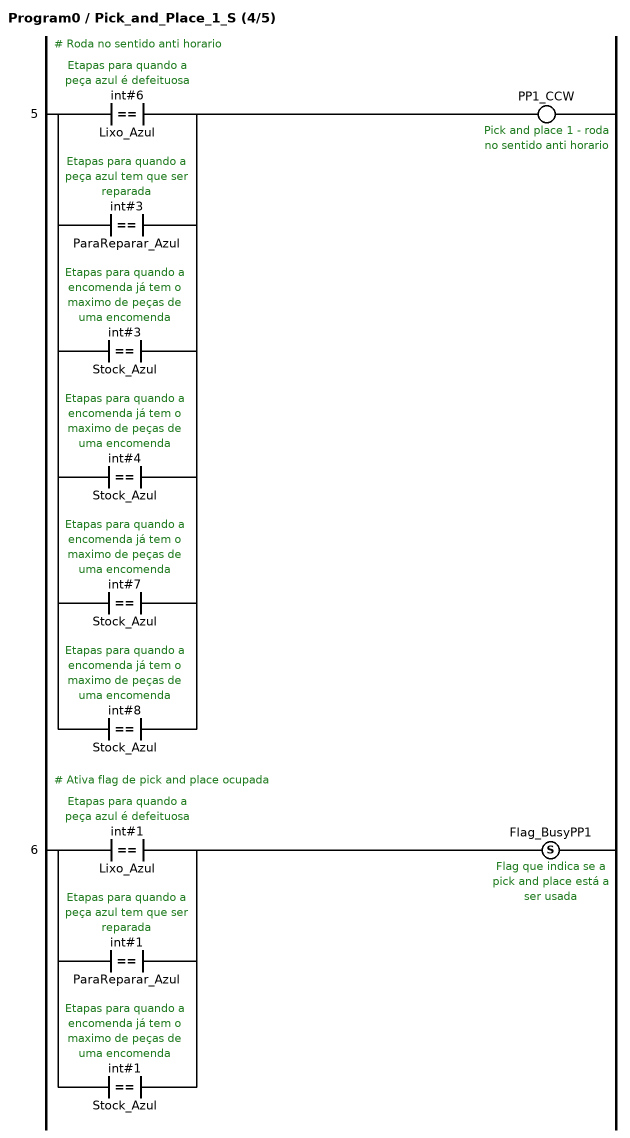
(* [picture p48: Program0 / Pick_and_Place_1_S, rungs 5-6] *)
(* Rung 5: # Roda no sentido anti horario *)
PP1_CCW := (int#6 = Lixo_Azul) OR (int#3 = ParaReparar_Azul) OR (int#3 = Stock_Azul) OR (int#4 = Stock_Azul) OR (int#7 = Stock_Azul) OR (int#8 = Stock_Azul);
(* Rung 6: # Ativa flag de pick and place ocupada *)
IF (int#1 = Lixo_Azul) OR (int#1 = ParaReparar_Azul) OR (int#1 = Stock_Azul) THEN
    Flag_BusyPP1 := TRUE;
END_IF;

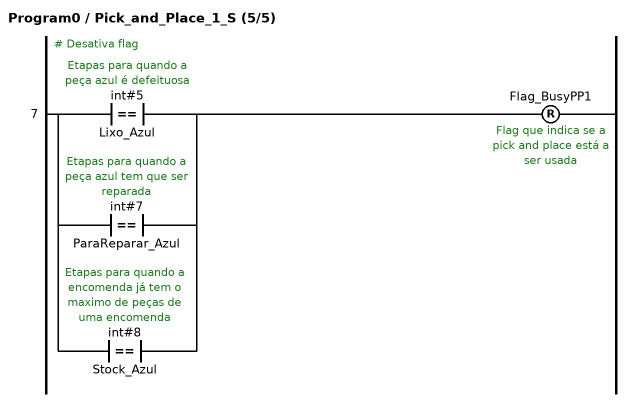
(* Rung 7: # Desativa flag *)
IF (int#5 = Lixo_Azul) OR (int#7 = ParaReparar_Azul) OR (int#8 = Stock_Azul) THEN
    Flag_BusyPP1 := FALSE;
END_IF;

(* Section Pick_and_Place_2_S: ladder, written here as Structured Text *)

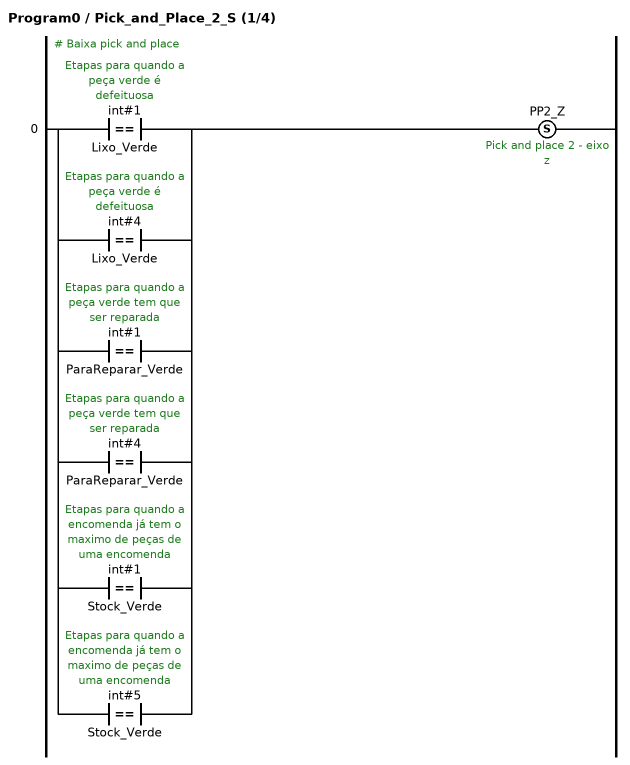
(* Rung 0: # Baixa pick and place *)
IF (int#1 = Lixo_Verde) OR (int#4 = Lixo_Verde) OR (int#1 = ParaReparar_Verde) OR (int#4 = ParaReparar_Verde) OR (int#1 = Stock_Verde) OR (int#5 = Stock_Verde) THEN
    PP2_Z := TRUE;
END_IF;

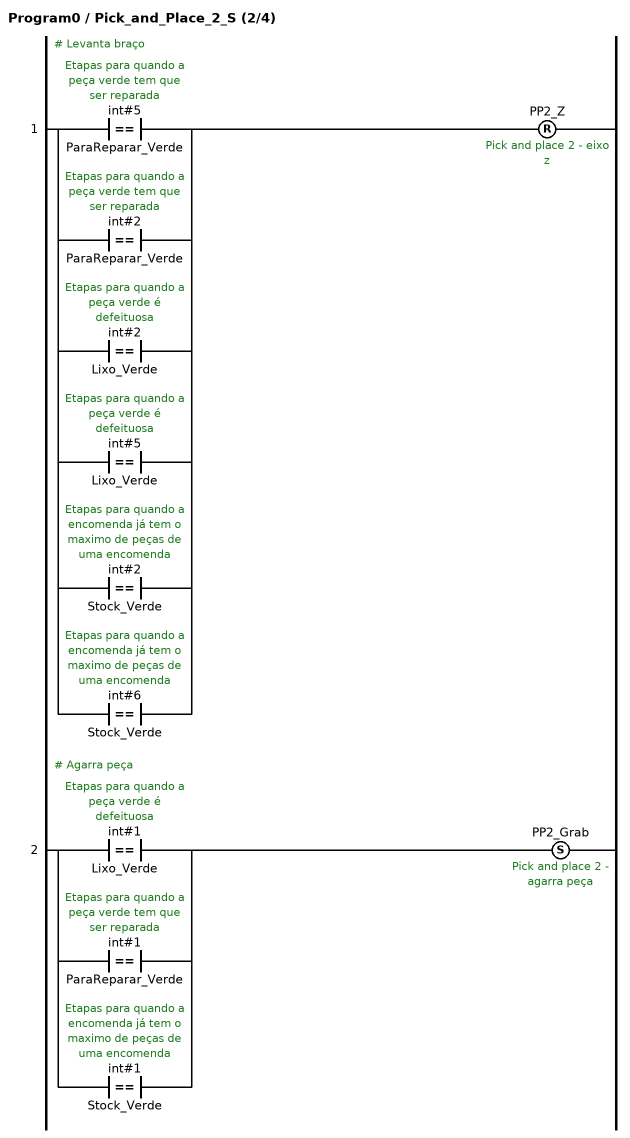
(* Rung 1: # Levanta braço *)
IF (int#5 = ParaReparar_Verde) OR (int#2 = ParaReparar_Verde) OR (int#2 = Lixo_Verde) OR (int#5 = Lixo_Verde) OR (int#2 = Stock_Verde) OR (int#6 = Stock_Verde) THEN
    PP2_Z := FALSE;
END_IF;
(* Rung 2: # Agarra peça *)
IF (int#1 = Lixo_Verde) OR (int#1 = ParaReparar_Verde) OR (int#1 = Stock_Verde) THEN
    PP2_Grab := TRUE;
END_IF;

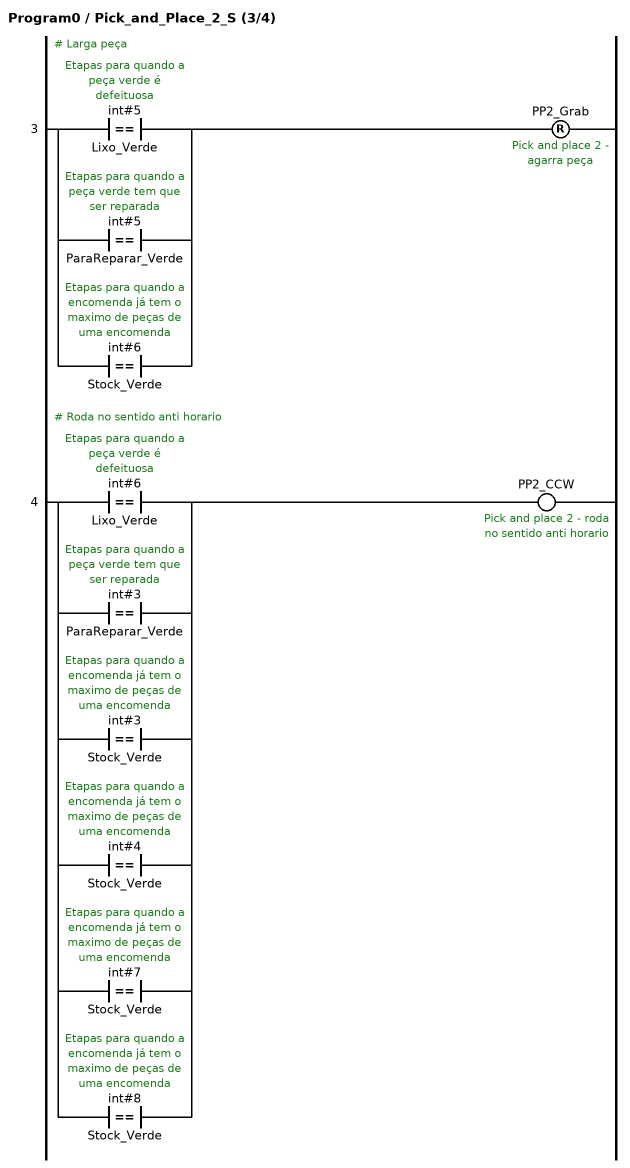
(* Rung 3: # Larga peça *)
IF (int#5 = Lixo_Verde) OR (int#5 = ParaReparar_Verde) OR (int#6 = Stock_Verde) THEN
    PP2_Grab := FALSE;
END_IF;
(* Rung 4: # Roda no sentido anti horario *)
PP2_CCW := (int#6 = Lixo_Verde) OR (int#3 = ParaReparar_Verde) OR (int#3 = Stock_Verde) OR (int#4 = Stock_Verde) OR (int#7 = Stock_Verde) OR (int#8 = Stock_Verde);

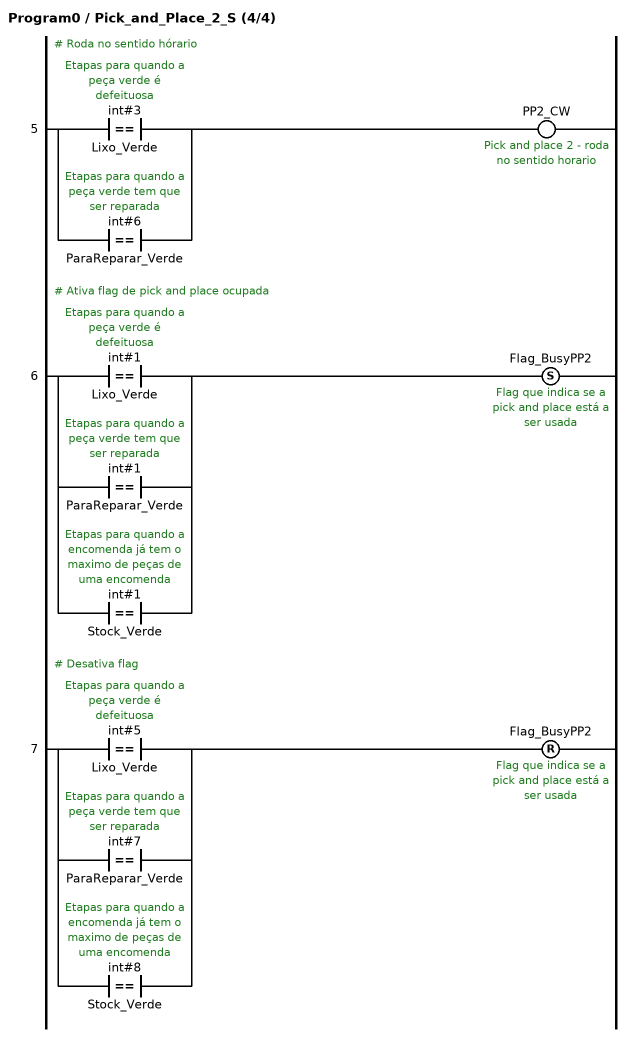
(* Rung 5: # Roda no sentido hórario *)
PP2_CW := (int#3 = Lixo_Verde) OR (int#6 = ParaReparar_Verde);
(* Rung 6: # Ativa flag de pick and place ocupada *)
IF (int#1 = Lixo_Verde) OR (int#1 = ParaReparar_Verde) OR (int#1 = Stock_Verde) THEN
    Flag_BusyPP2 := TRUE;
END_IF;
(* Rung 7: # Desativa flag *)
IF (int#5 = Lixo_Verde) OR (int#7 = ParaReparar_Verde) OR (int#8 = Stock_Verde) THEN
    Flag_BusyPP2 := FALSE;
END_IF;

(* Section Botoes: ladder, written here as Structured Text *)

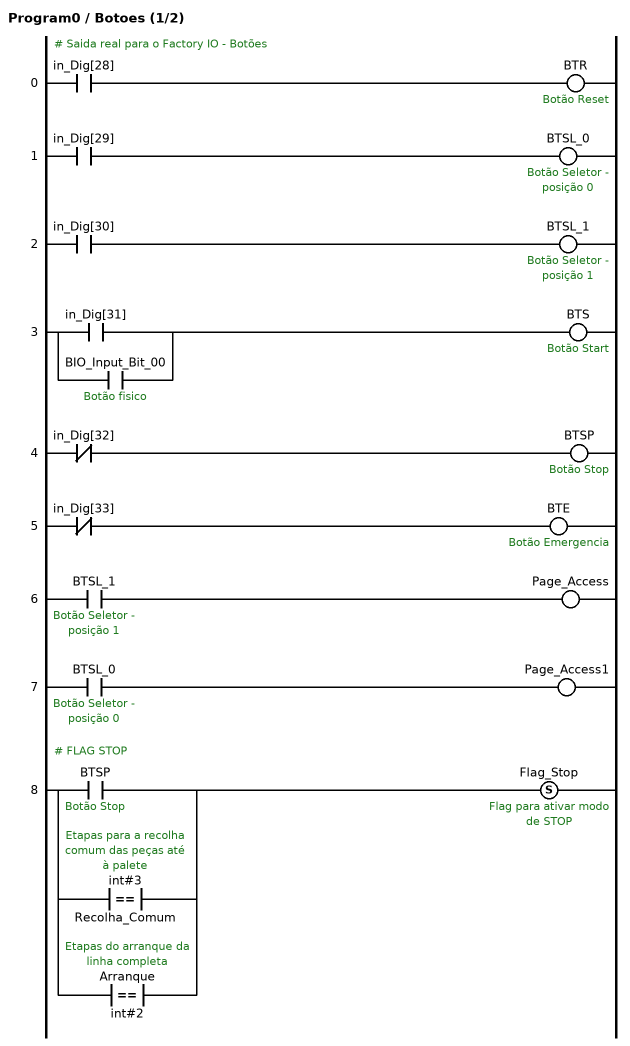
(* Rung 0: # Saida real para o Factory IO - Botões *)
BTR := in_Dig[28];
(* Rung 1 *)
BTSL_0 := in_Dig[29];
(* Rung 2 *)
BTSL_1 := in_Dig[30];
(* Rung 3 *)
BTS := in_Dig[31] OR BIO_Input_Bit_00;
(* Rung 4 *)
BTSP := NOT in_Dig[32];
(* Rung 5 *)
BTE := NOT in_Dig[33];
(* Rung 6 *)
Page_Access := BTSL_1;
(* Rung 7 *)
Page_Access1 := BTSL_0;
(* Rung 8: # FLAG STOP *)
IF BTSP OR (int#3 = Recolha_Comum) OR (Arranque = int#2) THEN Flag_Stop := TRUE; END_IF;

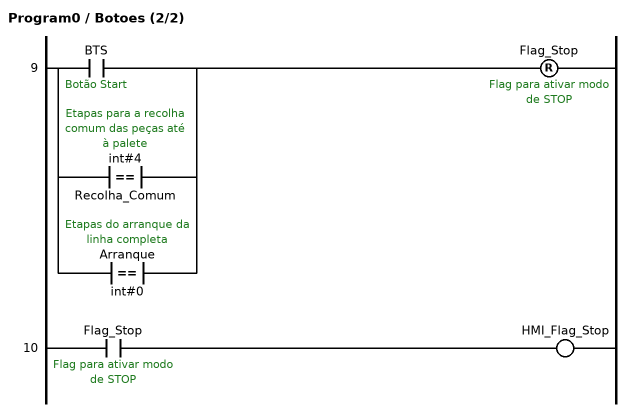
(* Rung 9 *)
IF BTS OR (int#4 = Recolha_Comum) OR (Arranque = int#0) THEN Flag_Stop := FALSE; END_IF;
(* Rung 10 *)
HMI_Flag_Stop := Flag_Stop;

(* Section Opto_Switches: ladder, written here as Structured Text *)

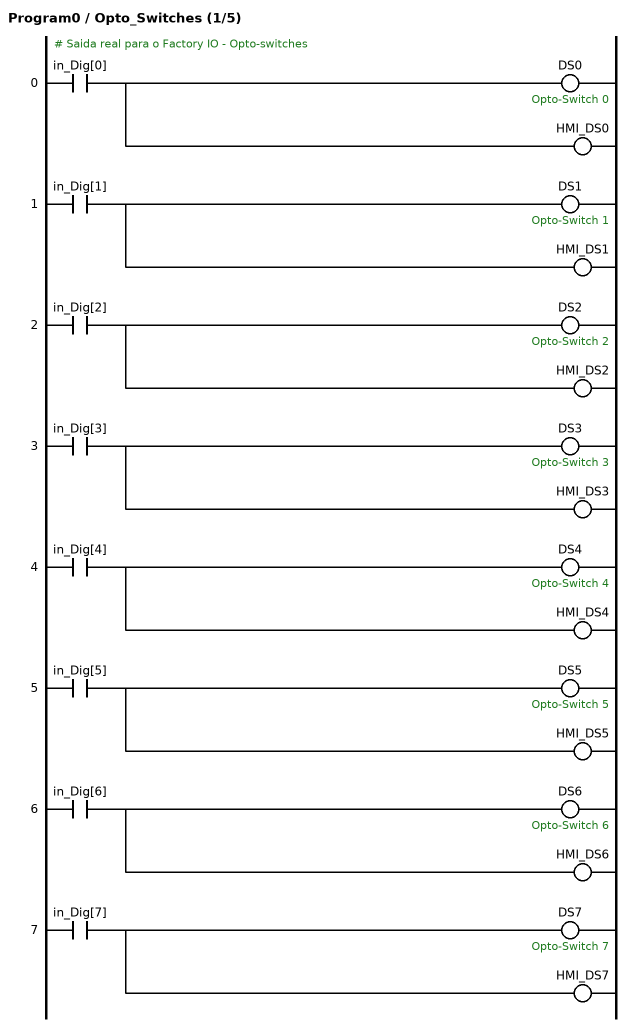
(* Rung 0: # Saida real para o Factory IO - Opto-switches *)
DS0 := in_Dig[0];
HMI_DS0 := in_Dig[0];
(* Rung 1 *)
DS1 := in_Dig[1];
HMI_DS1 := in_Dig[1];
(* Rung 2 *)
DS2 := in_Dig[2];
HMI_DS2 := in_Dig[2];
(* Rung 3 *)
DS3 := in_Dig[3];
HMI_DS3 := in_Dig[3];
(* Rung 4 *)
DS4 := in_Dig[4];
HMI_DS4 := in_Dig[4];
(* Rung 5 *)
DS5 := in_Dig[5];
HMI_DS5 := in_Dig[5];
(* Rung 6 *)
DS6 := in_Dig[6];
HMI_DS6 := in_Dig[6];
(* Rung 7 *)
DS7 := in_Dig[7];
HMI_DS7 := in_Dig[7];

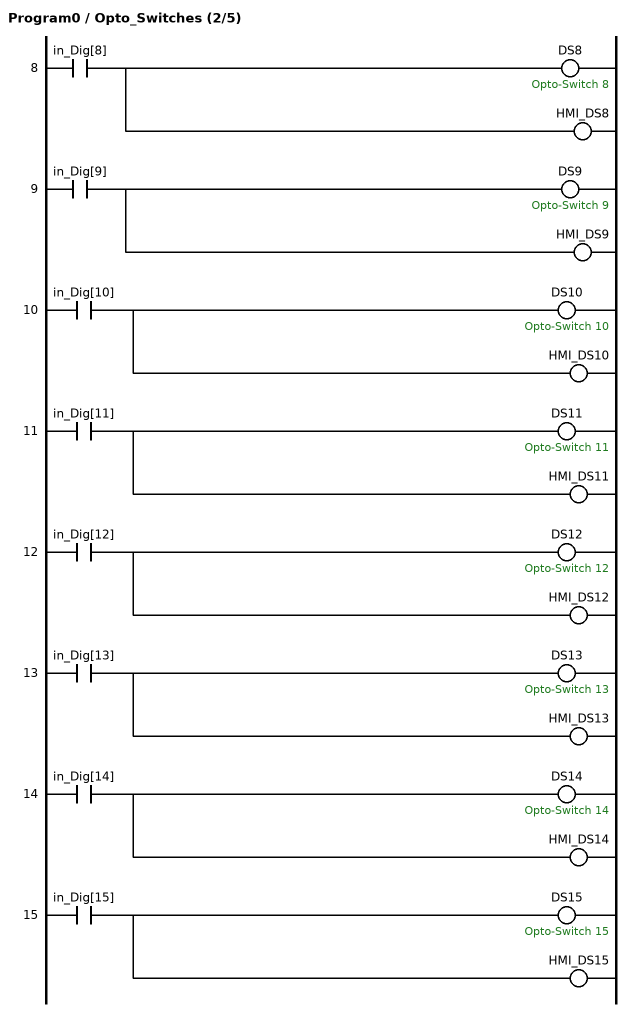
(* Rung 8 *)
DS8 := in_Dig[8];
HMI_DS8 := in_Dig[8];
(* Rung 9 *)
DS9 := in_Dig[9];
HMI_DS9 := in_Dig[9];
(* Rung 10 *)
DS10 := in_Dig[10];
HMI_DS10 := in_Dig[10];
(* Rung 11 *)
DS11 := in_Dig[11];
HMI_DS11 := in_Dig[11];
(* Rung 12 *)
DS12 := in_Dig[12];
HMI_DS12 := in_Dig[12];
(* Rung 13 *)
DS13 := in_Dig[13];
HMI_DS13 := in_Dig[13];
(* Rung 14 *)
DS14 := in_Dig[14];
HMI_DS14 := in_Dig[14];
(* Rung 15 *)
DS15 := in_Dig[15];
HMI_DS15 := in_Dig[15];

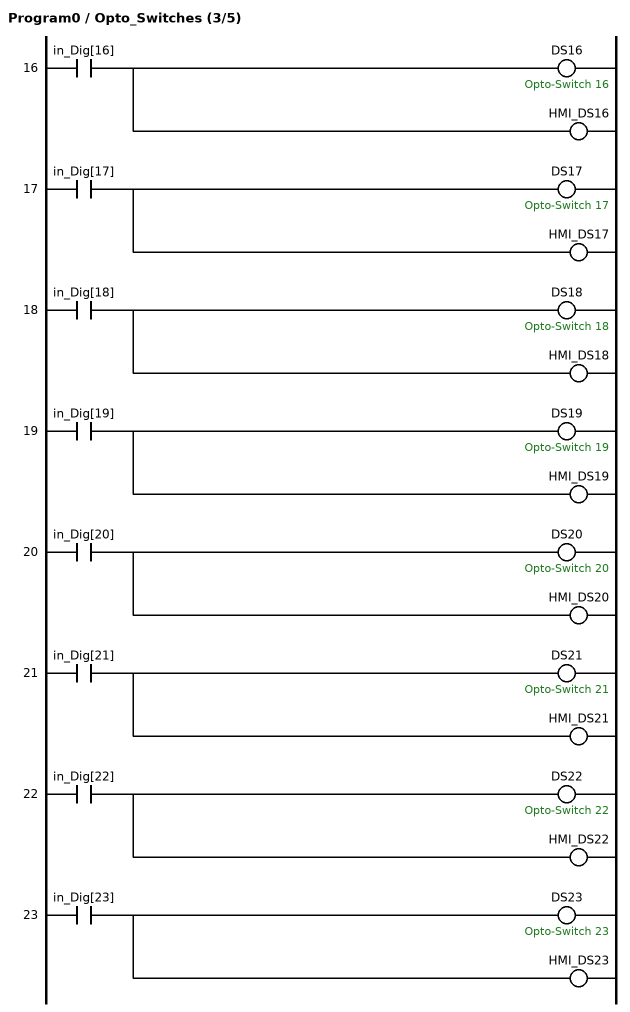
(* Rung 16 *)
DS16 := in_Dig[16];
HMI_DS16 := in_Dig[16];
(* Rung 17 *)
DS17 := in_Dig[17];
HMI_DS17 := in_Dig[17];
(* Rung 18 *)
DS18 := in_Dig[18];
HMI_DS18 := in_Dig[18];
(* Rung 19 *)
DS19 := in_Dig[19];
HMI_DS19 := in_Dig[19];
(* Rung 20 *)
DS20 := in_Dig[20];
HMI_DS20 := in_Dig[20];
(* Rung 21 *)
DS21 := in_Dig[21];
HMI_DS21 := in_Dig[21];
(* Rung 22 *)
DS22 := in_Dig[22];
HMI_DS22 := in_Dig[22];
(* Rung 23 *)
DS23 := in_Dig[23];
HMI_DS23 := in_Dig[23];

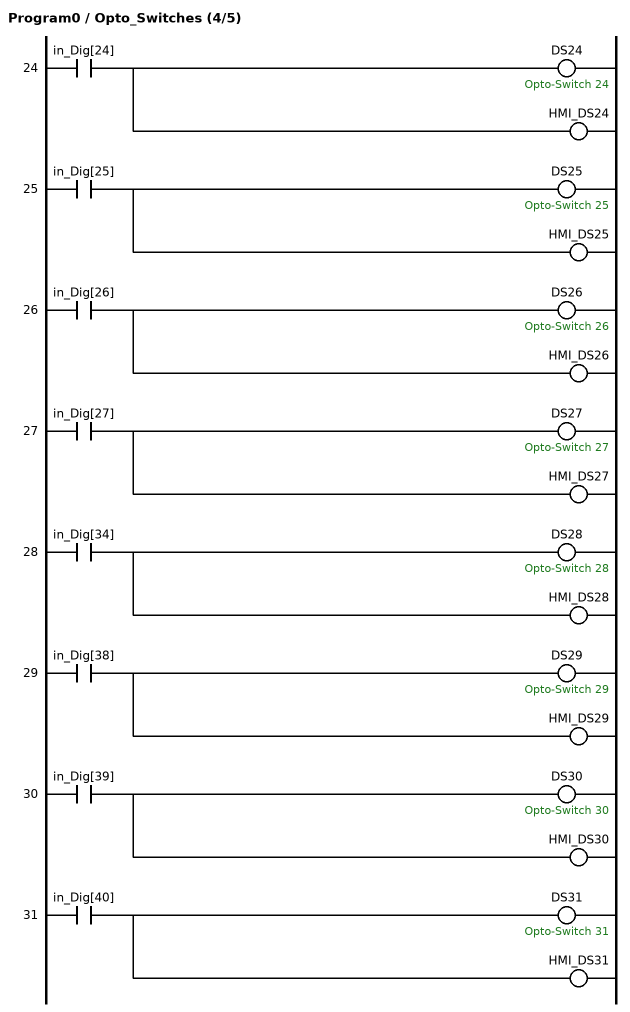
(* Rung 24 *)
DS24 := in_Dig[24];
HMI_DS24 := in_Dig[24];
(* Rung 25 *)
DS25 := in_Dig[25];
HMI_DS25 := in_Dig[25];
(* Rung 26 *)
DS26 := in_Dig[26];
HMI_DS26 := in_Dig[26];
(* Rung 27 *)
DS27 := in_Dig[27];
HMI_DS27 := in_Dig[27];
(* Rung 28 *)
DS28 := in_Dig[34];
HMI_DS28 := in_Dig[34];
(* Rung 29 *)
DS29 := in_Dig[38];
HMI_DS29 := in_Dig[38];
(* Rung 30 *)
DS30 := in_Dig[39];
HMI_DS30 := in_Dig[39];
(* Rung 31 *)
DS31 := in_Dig[40];
HMI_DS31 := in_Dig[40];

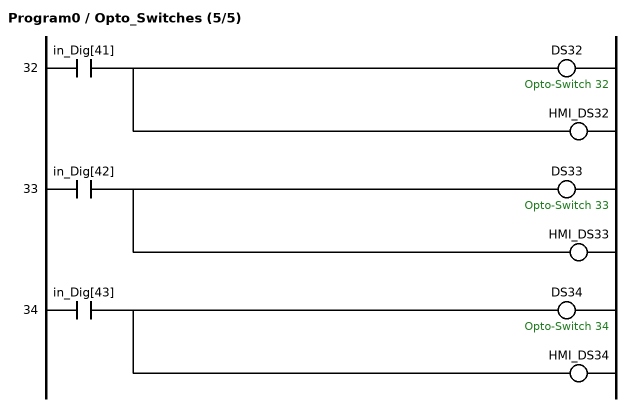
(* Rung 32 *)
DS32 := in_Dig[41];
HMI_DS32 := in_Dig[41];
(* Rung 33 *)
DS33 := in_Dig[42];
HMI_DS33 := in_Dig[42];
(* Rung 34 *)
DS34 := in_Dig[43];
HMI_DS34 := in_Dig[43];

(* Section Tapetes: ladder, written here as Structured Text *)

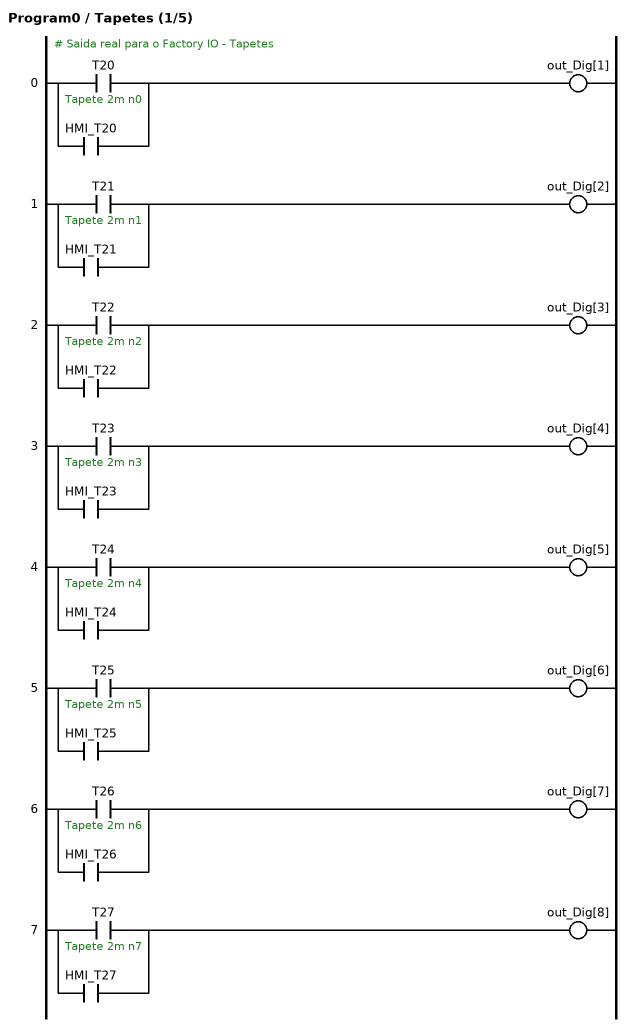
(* Rung 0: # Saida real para o Factory IO - Tapetes *)
out_Dig[1] := T20 OR HMI_T20;
(* Rung 1 *)
out_Dig[2] := T21 OR HMI_T21;
(* Rung 2 *)
out_Dig[3] := T22 OR HMI_T22;
(* Rung 3 *)
out_Dig[4] := T23 OR HMI_T23;
(* Rung 4 *)
out_Dig[5] := T24 OR HMI_T24;
(* Rung 5 *)
out_Dig[6] := T25 OR HMI_T25;
(* Rung 6 *)
out_Dig[7] := T26 OR HMI_T26;
(* Rung 7 *)
out_Dig[8] := T27 OR HMI_T27;

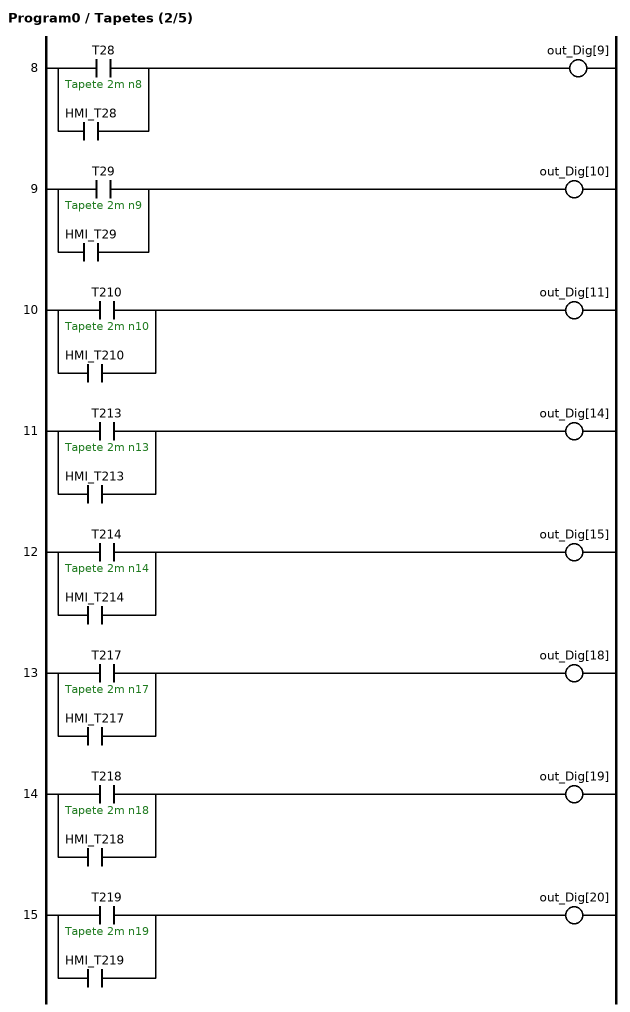
(* Rung 8 *)
out_Dig[9] := T28 OR HMI_T28;
(* Rung 9 *)
out_Dig[10] := T29 OR HMI_T29;
(* Rung 10 *)
out_Dig[11] := T210 OR HMI_T210;
(* Rung 11 *)
out_Dig[14] := T213 OR HMI_T213;
(* Rung 12 *)
out_Dig[15] := T214 OR HMI_T214;
(* Rung 13 *)
out_Dig[18] := T217 OR HMI_T217;
(* Rung 14 *)
out_Dig[19] := T218 OR HMI_T218;
(* Rung 15 *)
out_Dig[20] := T219 OR HMI_T219;

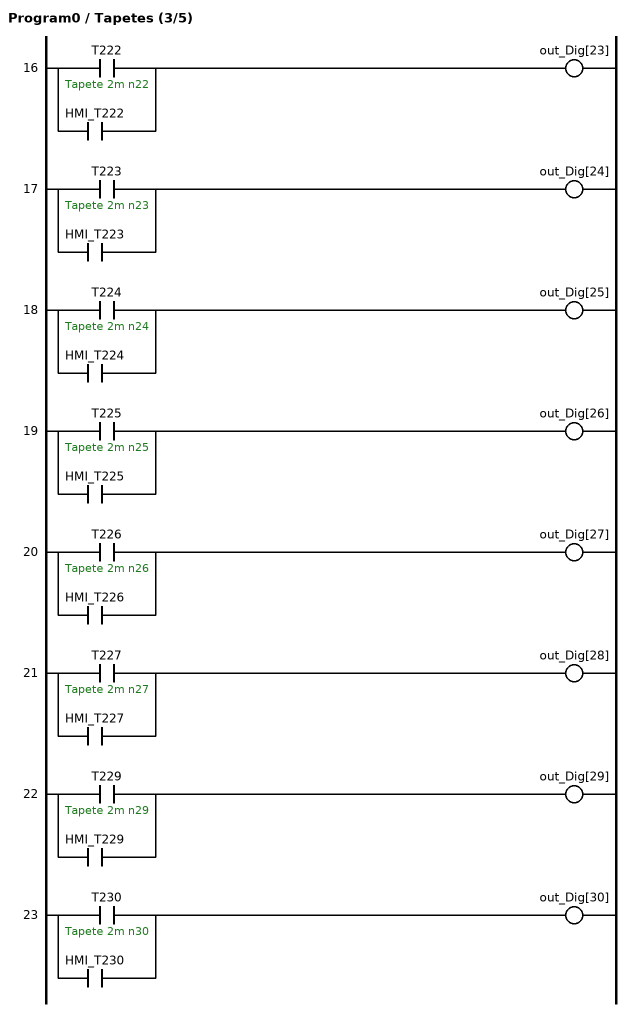
(* Rung 16 *)
out_Dig[23] := T222 OR HMI_T222;
(* Rung 17 *)
out_Dig[24] := T223 OR HMI_T223;
(* Rung 18 *)
out_Dig[25] := T224 OR HMI_T224;
(* Rung 19 *)
out_Dig[26] := T225 OR HMI_T225;
(* Rung 20 *)
out_Dig[27] := T226 OR HMI_T226;
(* Rung 21 *)
out_Dig[28] := T227 OR HMI_T227;
(* Rung 22 *)
out_Dig[29] := T229 OR HMI_T229;
(* Rung 23 *)
out_Dig[30] := T230 OR HMI_T230;

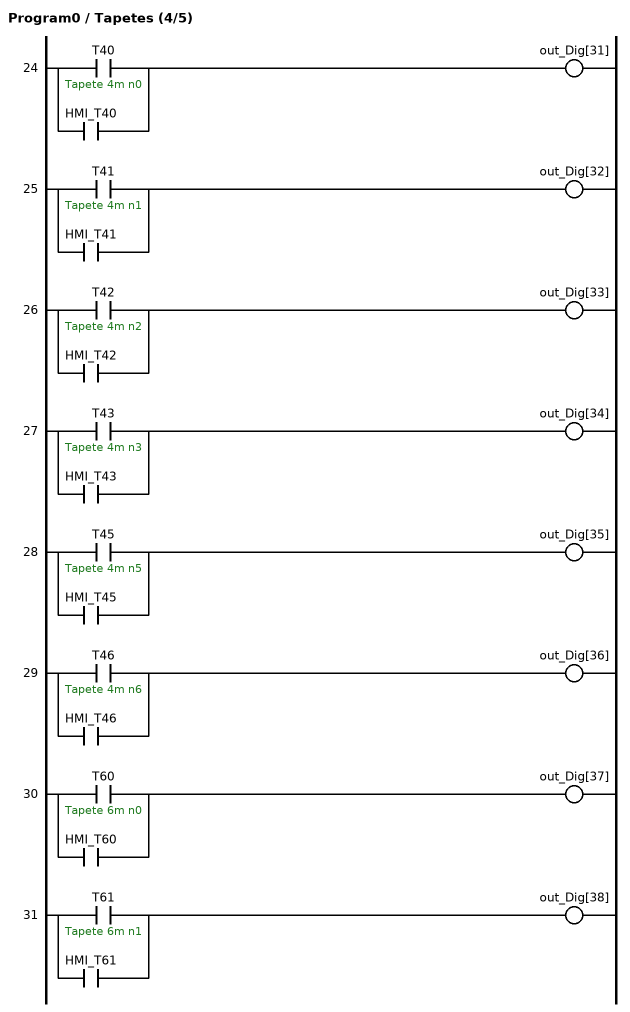
(* Rung 24 *)
out_Dig[31] := T40 OR HMI_T40;
(* Rung 25 *)
out_Dig[32] := T41 OR HMI_T41;
(* Rung 26 *)
out_Dig[33] := T42 OR HMI_T42;
(* Rung 27 *)
out_Dig[34] := T43 OR HMI_T43;
(* Rung 28 *)
out_Dig[35] := T45 OR HMI_T45;
(* Rung 29 *)
out_Dig[36] := T46 OR HMI_T46;
(* Rung 30 *)
out_Dig[37] := T60 OR HMI_T60;
(* Rung 31 *)
out_Dig[38] := T61 OR HMI_T61;

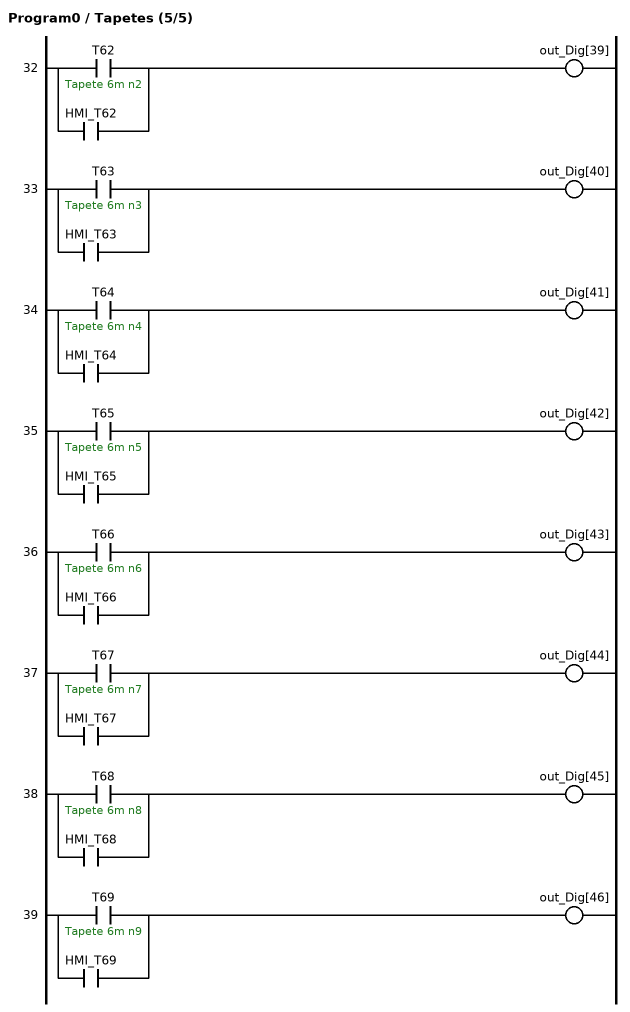
(* Rung 32 *)
out_Dig[39] := T62 OR HMI_T62;
(* Rung 33 *)
out_Dig[40] := T63 OR HMI_T63;
(* Rung 34 *)
out_Dig[41] := T64 OR HMI_T64;
(* Rung 35 *)
out_Dig[42] := T65 OR HMI_T65;
(* Rung 36 *)
out_Dig[43] := T66 OR HMI_T66;
(* Rung 37 *)
out_Dig[44] := T67 OR HMI_T67;
(* Rung 38 *)
out_Dig[45] := T68 OR HMI_T68;
(* Rung 39 *)
out_Dig[46] := T69 OR HMI_T69;

(* Section Tapetes_Analog: ladder, written here as Structured Text *)

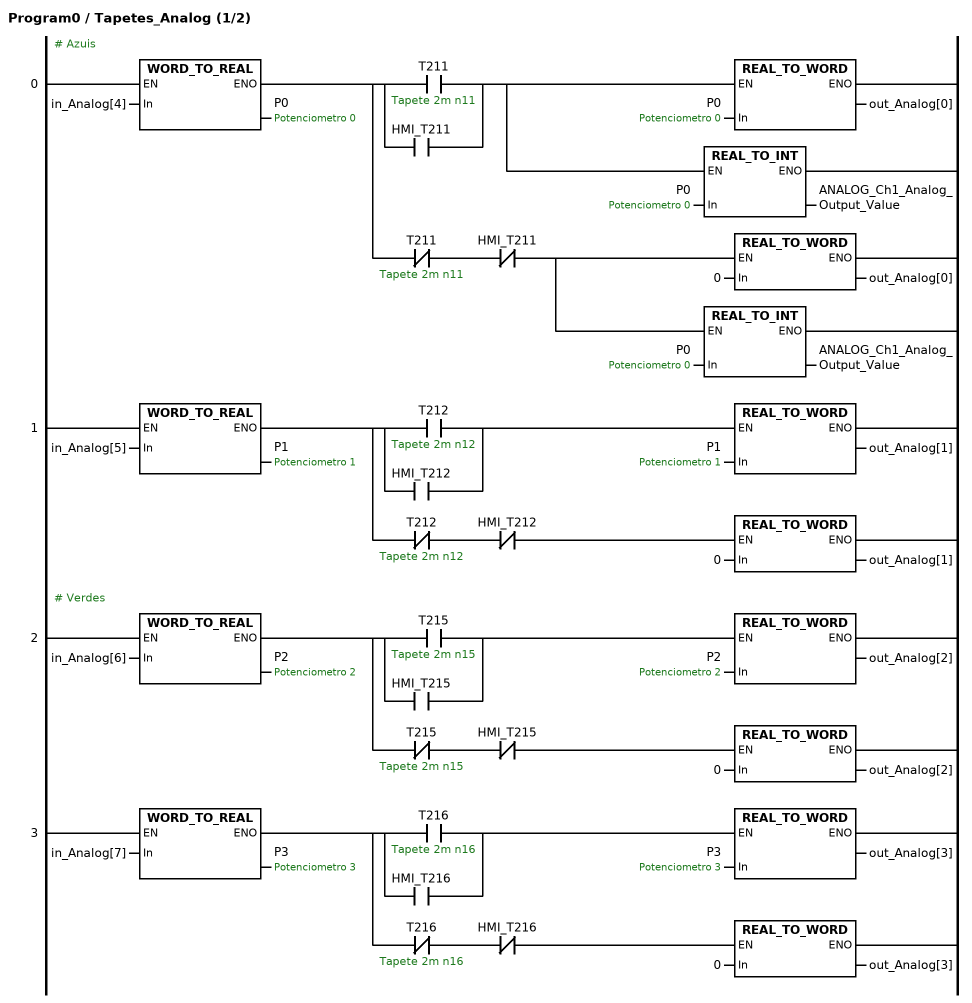
(* Rung 0: # Azuis *)
P0 := WORD_TO_REAL(In := in_Analog[4]);
IF T211 OR HMI_T211 THEN
    out_Analog[0] := REAL_TO_WORD(In := P0);
    ANALOG_Ch1_Analog_Output_Value := REAL_TO_INT(In := P0);
END_IF;
IF NOT T211 AND NOT HMI_T211 THEN
    out_Analog[0] := REAL_TO_WORD(In := 0);
    ANALOG_Ch1_Analog_Output_Value := REAL_TO_INT(In := P0);
END_IF;
(* Rung 1 *)
P1 := WORD_TO_REAL(In := in_Analog[5]);
IF T212 OR HMI_T212 THEN out_Analog[1] := REAL_TO_WORD(In := P1); END_IF;
IF NOT T212 AND NOT HMI_T212 THEN out_Analog[1] := REAL_TO_WORD(In := 0); END_IF;
(* Rung 2: # Verdes *)
P2 := WORD_TO_REAL(In := in_Analog[6]);
IF T215 OR HMI_T215 THEN out_Analog[2] := REAL_TO_WORD(In := P2); END_IF;
IF NOT T215 AND NOT HMI_T215 THEN out_Analog[2] := REAL_TO_WORD(In := 0); END_IF;
(* Rung 3 *)
P3 := WORD_TO_REAL(In := in_Analog[7]);
IF T216 OR HMI_T216 THEN out_Analog[3] := REAL_TO_WORD(In := P3); END_IF;
IF NOT T216 AND NOT HMI_T216 THEN out_Analog[3] := REAL_TO_WORD(In := 0); END_IF;

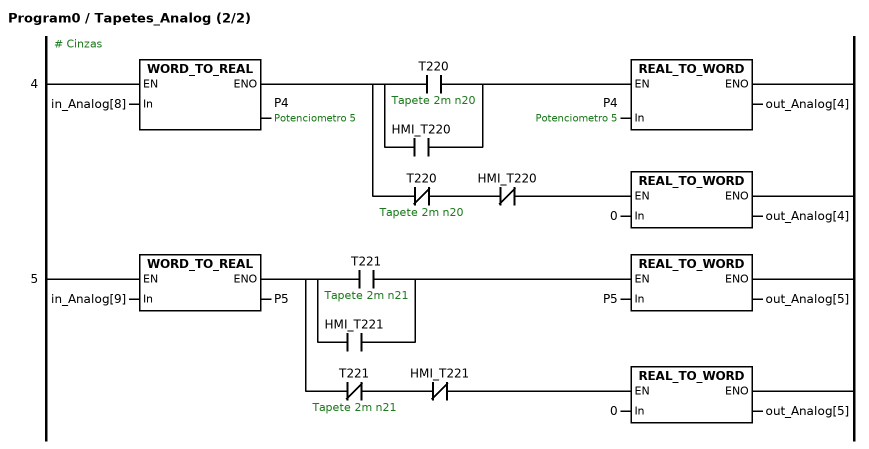
(* Rung 4: # Cinzas *)
P4 := WORD_TO_REAL(In := in_Analog[8]);
IF T220 OR HMI_T220 THEN out_Analog[4] := REAL_TO_WORD(In := P4); END_IF;
IF NOT T220 AND NOT HMI_T220 THEN out_Analog[4] := REAL_TO_WORD(In := 0); END_IF;
(* Rung 5 *)
P5 := WORD_TO_REAL(In := in_Analog[9]);
IF T221 OR HMI_T221 THEN out_Analog[5] := REAL_TO_WORD(In := P5); END_IF;
IF NOT T221 AND NOT HMI_T221 THEN out_Analog[5] := REAL_TO_WORD(In := 0); END_IF;

(* Section Tapetes_Curvos: ladder, written here as Structured Text *)

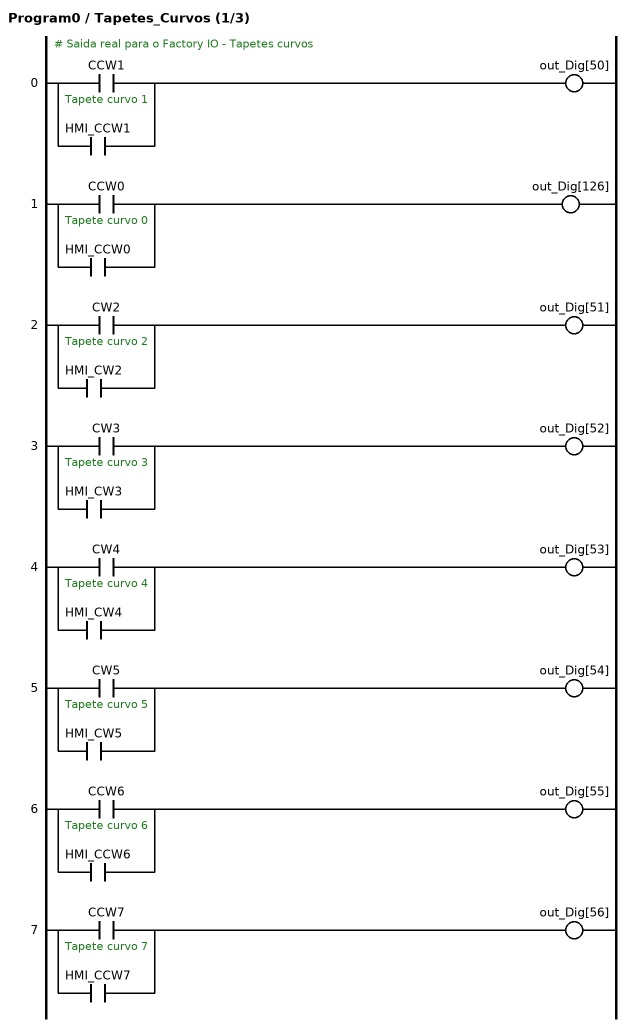
(* Rung 0: # Saida real para o Factory IO - Tapetes curvos *)
out_Dig[50] := CCW1 OR HMI_CCW1;
(* Rung 1 *)
out_Dig[126] := CCW0 OR HMI_CCW0;
(* Rung 2 *)
out_Dig[51] := CW2 OR HMI_CW2;
(* Rung 3 *)
out_Dig[52] := CW3 OR HMI_CW3;
(* Rung 4 *)
out_Dig[53] := CW4 OR HMI_CW4;
(* Rung 5 *)
out_Dig[54] := CW5 OR HMI_CW5;
(* Rung 6 *)
out_Dig[55] := CCW6 OR HMI_CCW6;
(* Rung 7 *)
out_Dig[56] := CCW7 OR HMI_CCW7;

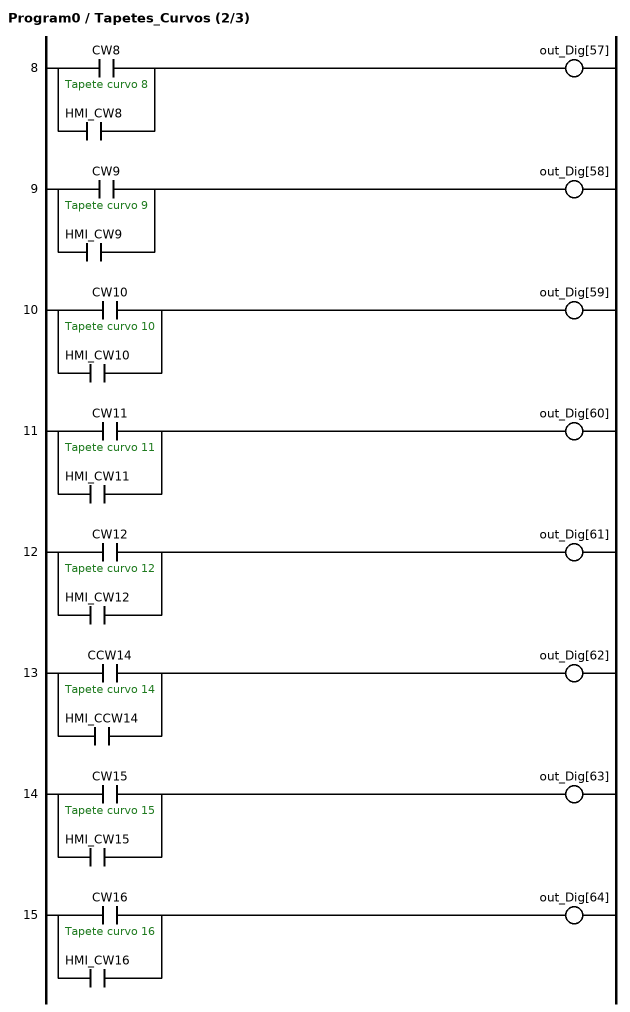
(* Rung 8 *)
out_Dig[57] := CW8 OR HMI_CW8;
(* Rung 9 *)
out_Dig[58] := CW9 OR HMI_CW9;
(* Rung 10 *)
out_Dig[59] := CW10 OR HMI_CW10;
(* Rung 11 *)
out_Dig[60] := CW11 OR HMI_CW11;
(* Rung 12 *)
out_Dig[61] := CW12 OR HMI_CW12;
(* Rung 13 *)
out_Dig[62] := CCW14 OR HMI_CCW14;
(* Rung 14 *)
out_Dig[63] := CW15 OR HMI_CW15;
(* Rung 15 *)
out_Dig[64] := CW16 OR HMI_CW16;

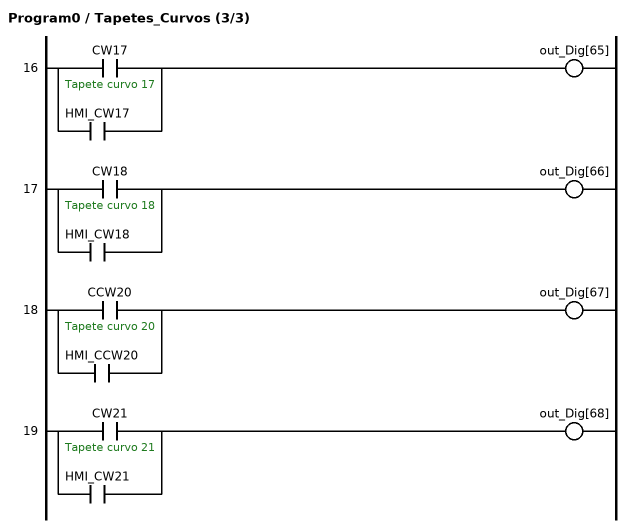
(* Rung 16 *)
out_Dig[65] := CW17 OR HMI_CW17;
(* Rung 17 *)
out_Dig[66] := CW18 OR HMI_CW18;
(* Rung 18 *)
out_Dig[67] := CCW20 OR HMI_CCW20;
(* Rung 19 *)
out_Dig[68] := CW21 OR HMI_CW21;

(* Section Pivot_Arms: ladder, written here as Structured Text *)

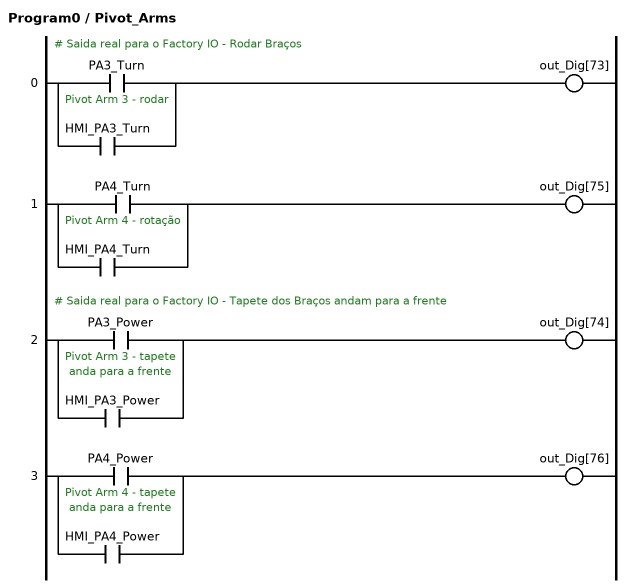
(* Rung 0: # Saida real para o Factory IO - Rodar Braços *)
out_Dig[73] := PA3_Turn OR HMI_PA3_Turn;
(* Rung 1 *)
out_Dig[75] := PA4_Turn OR HMI_PA4_Turn;
(* Rung 2: # Saida real para o Factory IO - Tapete dos Braços andam para a frente *)
out_Dig[74] := PA3_Power OR HMI_PA3_Power;
(* Rung 3 *)
out_Dig[76] := PA4_Power OR HMI_PA4_Power;

(* Section Balacas: ladder, written here as Structured Text *)

